TYPE "ST_CylinderParCfg"
VERSION : 0.1
   STRUCT
      SchemaVersion : UInt := 1;
      Timeout : Time := T#8S;
   END_STRUCT;

END_TYPE

